(* IEC 61131-3 sources: plc-vscode/tests/st/test-ready/trust-platform/examples/OSCAT/wind_speed_alarm/non-oop/src, 3 files *)

(* ---- Configuration.st ---- *)
CONFIGURATION WindSpeedAlarmClassicConfiguration
RESOURCE Cpu0 ON PLC
    TASK MainTask (INTERVAL := T#100ms, PRIORITY := 1);
    PROGRAM Main WITH MainTask : Main;
END_RESOURCE
END_CONFIGURATION

(* ---- Main.st ---- *)
PROGRAM Main
VAR
    WindAlarm : HYST;
    WindMetersPerSecond : REAL := REAL#10.0;
    BeaufortIndex : INT;
    AlarmActive : BOOL;
END_VAR

BeaufortIndex := MS_TO_BFT(MS := WindMetersPerSecond);
WindAlarm(In := WindMetersPerSecond, HIGH_LIMIT := REAL#8.0, LOW_LIMIT := REAL#3.0);
AlarmActive := WindAlarm.Q;
END_PROGRAM

(* ---- Tests.st ---- *)
TEST_PROGRAM WindSpeedAlarmClassicConvertsAndRaisesAlarm
VAR
    WindAlarm : HYST;
END_VAR

WindAlarm(In := REAL#10.0, HIGH_LIMIT := REAL#8.0, LOW_LIMIT := REAL#3.0);

ASSERT_EQUAL(EXPECTED := MS_TO_BFT(MS := REAL#10.0), ACTUAL := MS_TO_BFT(MS := REAL#10.0));
ASSERT_TRUE(IN := WindAlarm.Q);
END_TEST_PROGRAM
